TYPE ST_Machine_Command :
STRUCT
	Stop :BOOL;
END_STRUCT
END_TYPE

(* stored: Version 1.1.0.1, ProductVersion 3.1.4024.15
   DUT ST_Machine_Command: Id {4f6366d3-f1a2-4ca6-ae2b-7ab42fd8f7c1} *)
